// Core 3.10.2: deterministic typed walk, one bounded response window.
// Static facets carry no write capability. Every reused slot is cleared.
FUNCTION "FRK_ConfigRevision" : UDInt
{ S7_Optimized_Access := 'TRUE' }
VERSION : 0.1
VAR_INPUT
    Previous : UDInt;
END_VAR
VAR_TEMP
    Stamp : DTL;
    ResultCode : Int;
    Generation : ULInt;
END_VAR
BEGIN
    #FRK_ConfigRevision := #Previous + 1;
    #ResultCode := RD_SYS_T(OUT => #Stamp);
    IF #ResultCode = 0 THEN
        #Generation := LDT_TO_ULINT(DTL_TO_LDT(#Stamp)) / ULINT#1000000;
        #FRK_ConfigRevision := ULINT_TO_UDINT(#Generation MOD ULINT#4294967296);
    END_IF;
    IF #FRK_ConfigRevision = #Previous THEN #FRK_ConfigRevision := #Previous + 1; END_IF;
    IF #FRK_ConfigRevision = 0 THEN #FRK_ConfigRevision := 1; END_IF;
END_FUNCTION

FUNCTION "FRK_ConfigBegin" : Void
{ S7_Optimized_Access := 'TRUE' }
VERSION : 0.1
VAR_INPUT
    PageIndex : DInt;
    Revision : UDInt;
END_VAR
VAR_IN_OUT
    Cursor : "FRK_ConfigCursor";
    Page : "ST_ConfigPage";
END_VAR
VAR_TEMP
    Index : Int;
END_VAR
BEGIN
    #Cursor.Position := 0;
    #Cursor.First := 0;
    #Page.Revision := #Revision;
    #Page.PageIndex := 0;
    IF #PageIndex >= 0 AND #PageIndex <= 32767 THEN
        #Cursor.First := #PageIndex * 16;
        #Page.PageIndex := DINT_TO_INT(#PageIndex);
    END_IF;
    #Page.PageCount := 1;
    #Page.EntryCount := 0;
    "FRK_UnitScratch".EmptyConfigEntry.ValueType := 1;
    "FRK_UnitScratch".EmptyConfigEntry.Readable := TRUE;
    FOR #Index := 1 TO 16 DO
        #Page.Entries[#Index] := "FRK_UnitScratch".EmptyConfigEntry;
    END_FOR;
END_FUNCTION

FUNCTION "FRK_ConfigAppend" : Void
{ S7_Optimized_Access := 'TRUE' }
VERSION : 0.1
VAR_INPUT
    Scope : String;
    Item : String;
    ValueText : WString;
    ValueType : DInt;
    ReadLevel : DInt;
    Readable : Bool;
END_VAR
VAR_IN_OUT
    Cursor : "FRK_ConfigCursor";
    Page : "ST_ConfigPage";
END_VAR
VAR_TEMP
    Slot : DInt;
END_VAR
BEGIN
    #Slot := #Cursor.Position - #Cursor.First;
    #Cursor.Position := #Cursor.Position + 1;
    IF #Slot < 0 OR #Slot >= 16 THEN RETURN; END_IF;
    #Slot := #Slot + 1;
    #Page.Entries[#Slot].Scope := STRING_TO_WSTRING(#Scope);
    #Page.Entries[#Slot].Item := STRING_TO_WSTRING(#Item);
    #Page.Entries[#Slot].ValueType := #ValueType;
    #Page.Entries[#Slot].ReadLevel := #ReadLevel;
    #Page.Entries[#Slot].Readable := #Readable;
    IF #Readable THEN #Page.Entries[#Slot].ValueText := #ValueText; END_IF;
    #Page.EntryCount := DINT_TO_INT(#Slot);
END_FUNCTION

FUNCTION "FRK_ConfigFinish" : Void
{ S7_Optimized_Access := 'TRUE' }
VERSION : 0.1
VAR_IN_OUT
    Cursor : "FRK_ConfigCursor";
    Page : "ST_ConfigPage";
END_VAR
BEGIN
    #Page.PageCount := DINT_TO_INT((#Cursor.Position + 16 - 1) / 16);
    IF #Page.PageCount < 1 THEN #Page.PageCount := 1; END_IF;
END_FUNCTION

FUNCTION "FRK_ConfigCatalog" : Void
{ S7_Optimized_Access := 'TRUE' }
VERSION : 0.1
VAR_INPUT
    Scope : String;
    Count : Int;
    Catalog : Array[1..12] of "ST_CommandInfo";
    ReadLevel : DInt;
    Readable : Bool;
END_VAR
VAR_IN_OUT
    Cursor : "FRK_ConfigCursor";
    Page : "ST_ConfigPage";
END_VAR
VAR_TEMP
    Index : Int;
    IndexText : String[8];
    Prefix : String[254];
    Item : String[254];
END_VAR
BEGIN
    "FRK_ConfigAppend"(Scope := #Scope, Item := 'CatalogCount', ValueText := STRING_TO_WSTRING(INT_TO_STRING(#Count)), ValueType := 0, ReadLevel := #ReadLevel, Readable := #Readable, Cursor := #Cursor, Page := #Page);
    FOR #Index := 1 TO #Count DO
        IF #Index > 12 THEN EXIT; END_IF;
        #IndexText := INT_TO_STRING(#Index);
        IF #IndexText[1] = '+' THEN #IndexText := DELETE(IN := #IndexText, L := 1, P := 1); END_IF;
        #Prefix := CONCAT(IN1 := 'Catalog/Catalog[', IN2 := #IndexText);
        #Prefix := CONCAT(IN1 := #Prefix, IN2 := ']/');
        #Item := CONCAT(IN1 := #Prefix, IN2 := 'Value');
        "FRK_ConfigAppend"(Scope := #Scope, Item := #Item, ValueText := STRING_TO_WSTRING(DINT_TO_STRING(#Catalog[#Index].Value)), ValueType := 0, ReadLevel := #ReadLevel, Readable := #Readable, Cursor := #Cursor, Page := #Page);
        #Item := CONCAT(IN1 := #Prefix, IN2 := 'Label');
        "FRK_ConfigAppend"(Scope := #Scope, Item := #Item, ValueText := STRING_TO_WSTRING(#Catalog[#Index].Label), ValueType := 1, ReadLevel := #ReadLevel, Readable := #Readable, Cursor := #Cursor, Page := #Page);
        #Item := CONCAT(IN1 := #Prefix, IN2 := 'Style');
        "FRK_ConfigAppend"(Scope := #Scope, Item := #Item, ValueText := STRING_TO_WSTRING(DINT_TO_STRING(#Catalog[#Index].Style)), ValueType := 0, ReadLevel := #ReadLevel, Readable := #Readable, Cursor := #Cursor, Page := #Page);
    END_FOR;
END_FUNCTION

FUNCTION "FRK_ConfigUnit" : Void
{ S7_Optimized_Access := 'TRUE' }
VERSION : 0.1
VAR_INPUT
    Scope : String;
    Policy : Array[0..6] of "ST_ModePolicy";
    ModelCount : Int;
    ReadLevel : DInt;
    Readable : Bool;
END_VAR
VAR_IN_OUT
    Cursor : "FRK_ConfigCursor";
    Page : "ST_ConfigPage";
END_VAR
VAR_TEMP
    Index : Int;
    IndexText : String[8];
    Prefix : String[254];
    Item : String[254];
END_VAR
BEGIN
    "FRK_ConfigAppend"(Scope := #Scope, Item := 'CatalogCount', ValueText := WSTRING#'0', ValueType := 0, ReadLevel := #ReadLevel, Readable := #Readable, Cursor := #Cursor, Page := #Page);
    "FRK_ConfigAppend"(Scope := #Scope, Item := 'AvailableModelCount', ValueText := INT_TO_WSTRING(#ModelCount), ValueType := 0, ReadLevel := #ReadLevel, Readable := #Readable, Cursor := #Cursor, Page := #Page);
    FOR #Index := 0 TO 6 DO
        #IndexText := INT_TO_STRING(#Index);
        IF #IndexText[1] = '+' THEN #IndexText := DELETE(IN := #IndexText, L := 1, P := 1); END_IF;
        #Prefix := CONCAT(IN1 := 'ModePolicy/ModePolicy[', IN2 := #IndexText);
        #Prefix := CONCAT(IN1 := #Prefix, IN2 := ']/');
        #Item := CONCAT(IN1 := #Prefix, IN2 := 'Shield');
        "FRK_ConfigAppend"(Scope := #Scope, Item := #Item, ValueText := STRING_TO_WSTRING(DINT_TO_STRING(#Policy[#Index].Shield)), ValueType := 0, ReadLevel := #ReadLevel, Readable := #Readable, Cursor := #Cursor, Page := #Page);
        #Item := CONCAT(IN1 := #Prefix, IN2 := 'Style');
        "FRK_ConfigAppend"(Scope := #Scope, Item := #Item, ValueText := STRING_TO_WSTRING(DINT_TO_STRING(#Policy[#Index].Style)), ValueType := 0, ReadLevel := #ReadLevel, Readable := #Readable, Cursor := #Cursor, Page := #Page);
    END_FOR;
END_FUNCTION

// Core 8.3: one owning active list / closed ring, with optional event callback.
FUNCTION "FRK_AlarmNotify" : Void
{ S7_Optimized_Access := 'TRUE' }
VERSION : 0.1
VAR_INPUT
    Ev : "ST_AlarmEvent";
END_VAR
VAR_IN_OUT
    AlarmLog : "FRK_AlarmLog";
END_VAR
BEGIN
    RETURN; // No event sink supplied by the composition declaration.
END_FUNCTION

FUNCTION "FRK_AlarmRefresh" : Void
{ S7_Optimized_Access := 'TRUE' }
VERSION : 0.1
VAR_IN_OUT
    AlarmLog : "FRK_AlarmLog";
END_VAR
VAR_TEMP
    Index : Int;
END_VAR
BEGIN
    #AlarmLog.NActive := 0;
    #AlarmLog.Blocking := FALSE;
    FOR #Index := 1 TO 16 DO
        IF #AlarmLog.Active[#Index].State <> 0 THEN
            #AlarmLog.NActive := #AlarmLog.NActive + 1;
            IF #AlarmLog.Active[#Index].ResetClass = 1 THEN #AlarmLog.Blocking := TRUE; END_IF;
        END_IF;
    END_FOR;
END_FUNCTION

FUNCTION "FRK_AlarmBegin" : Void
{ S7_Optimized_Access := 'TRUE' }
VERSION : 0.1
VAR_INPUT
    Startup : Bool;
END_VAR
VAR_IN_OUT
    AlarmLog : "FRK_AlarmLog";
END_VAR
VAR_TEMP
    Index : Int;
END_VAR
BEGIN
    FOR #Index := 1 TO 16 DO
        #AlarmLog.Touched[#Index] := FALSE;
        IF #Startup THEN
            #AlarmLog.Active[#Index] := "FRK_UnitScratch".EmptyEvent;
            #AlarmLog.Automatic[#Index] := FALSE;
            #AlarmLog.ComeMs[#Index] := 0;
        END_IF;
    END_FOR;
    IF #Startup THEN
        FOR #Index := 1 TO 64 DO #AlarmLog.Ring[#Index] := "FRK_UnitScratch".EmptyEvent; END_FOR;
        #AlarmLog.RingHead := 0;
        #AlarmLog.RingUsed := 0;
        #AlarmLog.Truncated := FALSE;
    END_IF;
    "FRK_AlarmRefresh"(AlarmLog := #AlarmLog);
END_FUNCTION

FUNCTION "FRK_AlarmRaise" : Int
{ S7_Optimized_Access := 'TRUE' }
VERSION : 0.1
VAR_INPUT
    Diag : "ST_Diagnostic";
    ResetClass : DInt;
END_VAR
VAR_IN_OUT
    AlarmLog : "FRK_AlarmLog";
END_VAR
VAR_TEMP
    Slot : Int;
    Stamp : DTL;
    ResultCode : Int;
    Rational : "ST_Diagnostic";
END_VAR
BEGIN
    #FRK_AlarmRaise := 0;
    IF #ResetClass < 0 OR #ResetClass > 1
        OR #Diag.Severity < 0 OR #Diag.Severity > 2
        OR #Diag.Category < 0 OR #Diag.Category > 2
        OR #Diag.SourcePath = WSTRING#'' OR #Diag.Description = WSTRING#'' THEN RETURN; END_IF;
    FOR #Slot := 1 TO 16 DO
        IF #AlarmLog.Active[#Slot].State = 0 THEN
            #Rational := #Diag;
            "FRK_Rationalize"(Diag := #Rational);
            #AlarmLog.Active[#Slot] := "FRK_UnitScratch".EmptyEvent;
            #AlarmLog.Active[#Slot].ReasonCode := #Rational.ReasonCode;
            #AlarmLog.Active[#Slot].Description := #Rational.Description;
            #AlarmLog.Active[#Slot].SourcePath := #Rational.SourcePath;
            #AlarmLog.Active[#Slot].IoTag := #Rational.IoTag;
            #AlarmLog.Active[#Slot].IoAddress := #Rational.IoAddress;
            #AlarmLog.Active[#Slot].Severity := #Rational.Severity;
            #AlarmLog.Active[#Slot].Category := #Rational.Category;
            #AlarmLog.Active[#Slot].ResetClass := #ResetClass;
            #AlarmLog.Active[#Slot].State := 1;
            #AlarmLog.ComeMs[#Slot] := "FRK_Clock".NowMs;
            #AlarmLog.Automatic[#Slot] := FALSE;
            #AlarmLog.Touched[#Slot] := FALSE;
            #ResultCode := RD_SYS_T(OUT => #Stamp);
            IF #ResultCode = 0 THEN #AlarmLog.Active[#Slot].ComeAt := DTL_TO_LDT(#Stamp); END_IF;
            // The UTC source has no proven synchronization witness yet.
            #AlarmLog.Active[#Slot].ComeTimeSynchronized := FALSE;
            "FRK_AlarmRefresh"(AlarmLog := #AlarmLog);
            "FRK_AlarmNotify"(AlarmLog := #AlarmLog, Ev := #AlarmLog.Active[#Slot]);
            #FRK_AlarmRaise := #Slot;
            RETURN;
        END_IF;
    END_FOR;
    #AlarmLog.Truncated := TRUE;
END_FUNCTION

FUNCTION "FRK_AlarmClose" : Void
{ S7_Optimized_Access := 'TRUE' }
VERSION : 0.1
VAR_INPUT
    Slot : Int;
END_VAR
VAR_IN_OUT
    AlarmLog : "FRK_AlarmLog";
END_VAR
BEGIN
    IF #Slot < 1 OR #Slot > 16 THEN RETURN; END_IF;
    IF #AlarmLog.Active[#Slot].State = 0 THEN RETURN; END_IF;
    #AlarmLog.Active[#Slot].State := 0;
    IF #AlarmLog.RingHead < 0 OR #AlarmLog.RingHead > 64 THEN #AlarmLog.RingHead := 0; END_IF;
    #AlarmLog.RingHead := (#AlarmLog.RingHead MOD 64) + 1;
    IF #AlarmLog.RingUsed >= 64 THEN #AlarmLog.Truncated := TRUE;
    ELSE #AlarmLog.RingUsed := #AlarmLog.RingUsed + 1; END_IF;
    #AlarmLog.Ring[#AlarmLog.RingHead] := #AlarmLog.Active[#Slot];
    #AlarmLog.Automatic[#Slot] := FALSE;
    "FRK_AlarmRefresh"(AlarmLog := #AlarmLog);
    "FRK_AlarmNotify"(AlarmLog := #AlarmLog, Ev := #AlarmLog.Ring[#AlarmLog.RingHead]);
END_FUNCTION

FUNCTION "FRK_AlarmGone" : Bool
{ S7_Optimized_Access := 'TRUE' }
VERSION : 0.1
VAR_INPUT
    Slot : Int;
END_VAR
VAR_IN_OUT
    AlarmLog : "FRK_AlarmLog";
END_VAR
VAR_TEMP
    Span : UDInt;
    Stamp : DTL;
    ResultCode : Int;
END_VAR
BEGIN
    #FRK_AlarmGone := FALSE;
    IF #Slot < 1 OR #Slot > 16 THEN RETURN; END_IF;
    IF #AlarmLog.Active[#Slot].State <> 1 THEN RETURN; END_IF;
    #ResultCode := RD_SYS_T(OUT => #Stamp);
    IF #ResultCode = 0 THEN #AlarmLog.Active[#Slot].GoneAt := DTL_TO_LDT(#Stamp); END_IF;
    #AlarmLog.Active[#Slot].GoneTimeSynchronized := FALSE;
    #Span := "FRK_Elapsed"(NewMs := "FRK_Clock".NowMs, OldMs := #AlarmLog.ComeMs[#Slot]);
    IF #Span > 2147483647 THEN #Span := 2147483647; END_IF;
    #AlarmLog.Active[#Slot].Duration := DINT_TO_TIME(UDINT_TO_DINT(#Span));
    IF #AlarmLog.Active[#Slot].ResetClass = 0 THEN
        "FRK_AlarmClose"(AlarmLog := #AlarmLog, Slot := #Slot);
    ELSE
        #AlarmLog.Active[#Slot].State := 2;
        #AlarmLog.Automatic[#Slot] := FALSE;
    END_IF;
    #FRK_AlarmGone := TRUE;
END_FUNCTION

FUNCTION "FRK_AlarmOperatorReset" : Void
{ S7_Optimized_Access := 'TRUE' }
VERSION : 0.1
VAR_IN_OUT
    AlarmLog : "FRK_AlarmLog";
END_VAR
VAR_TEMP
    Slot : Int;
    Gone : Bool;
    Stamp : DTL;
    ResultCode : Int;
END_VAR
BEGIN
    FOR #Slot := 1 TO 16 DO
        IF #AlarmLog.Active[#Slot].State <> 0 AND #AlarmLog.Active[#Slot].ResetClass = 1 THEN
            IF #AlarmLog.Active[#Slot].State = 1 THEN #Gone := "FRK_AlarmGone"(AlarmLog := #AlarmLog, Slot := #Slot); END_IF;
            #ResultCode := RD_SYS_T(OUT => #Stamp);
            IF #ResultCode = 0 THEN #AlarmLog.Active[#Slot].ResetAt := DTL_TO_LDT(#Stamp); END_IF;
            #AlarmLog.Active[#Slot].ResetTimeSynchronized := FALSE;
            "FRK_AlarmClose"(AlarmLog := #AlarmLog, Slot := #Slot);
        END_IF;
    END_FOR;
END_FUNCTION

FUNCTION "FRK_AlarmMessage" : Void
{ S7_Optimized_Access := 'TRUE' }
VERSION : 0.1
VAR_INPUT
    Reason : DInt;
    Description : WString;
    SourcePath : WString;
END_VAR
VAR_IN_OUT
    AlarmLog : "FRK_AlarmLog";
END_VAR
VAR_TEMP
    Diag : "ST_Diagnostic";
    Slot : Int;
    Gone : Bool;
END_VAR
BEGIN
    #Diag := "FRK_UnitScratch".EmptyDiagnostic;
    #Diag.ReasonCode := #Reason;
    #Diag.Description := #Description;
    #Diag.SourcePath := #SourcePath;
    #Diag.Severity := 0;
    #Diag.Category := 2;
    #Slot := "FRK_AlarmRaise"(AlarmLog := #AlarmLog, Diag := #Diag, ResetClass := 0);
    IF #Slot > 0 THEN #Gone := "FRK_AlarmGone"(AlarmLog := #AlarmLog, Slot := #Slot); END_IF;
END_FUNCTION

FUNCTION "FRK_AlarmCapture" : Void
{ S7_Optimized_Access := 'TRUE' }
VERSION : 0.1
VAR_IN_OUT
    AlarmLog : "FRK_AlarmLog";
    Core : "FRK_Core";
    Status : "ST_ModuleStatus";
END_VAR
VAR_TEMP
    Slot : Int;
END_VAR
BEGIN
    #Slot := #Core.FaultSlot;
    IF #Slot < 1 OR #Slot > 16 THEN #Slot := 0;
    ELSIF NOT #AlarmLog.Automatic[#Slot] OR #AlarmLog.Active[#Slot].State <> 1
        OR #AlarmLog.Active[#Slot].SourcePath <> #Status.Diagnostic.SourcePath
        OR #AlarmLog.Active[#Slot].ReasonCode <> #Status.Diagnostic.ReasonCode
        OR #AlarmLog.Active[#Slot].Description <> #Status.Diagnostic.Description THEN #Slot := 0; END_IF;
    IF #Core.Exec = 3 THEN
        IF #Slot = 0 THEN
            // Adopted first-outs share one active occurrence within this log.
            FOR #Slot := 1 TO 16 DO
                IF #AlarmLog.Automatic[#Slot] AND #AlarmLog.Active[#Slot].State = 1
                    AND #AlarmLog.Active[#Slot].SourcePath = #Status.Diagnostic.SourcePath
                    AND #AlarmLog.Active[#Slot].ReasonCode = #Status.Diagnostic.ReasonCode
                    AND #AlarmLog.Active[#Slot].Description = #Status.Diagnostic.Description THEN EXIT; END_IF;
            END_FOR;
            IF #Slot > 16 THEN #Slot := "FRK_AlarmRaise"(AlarmLog := #AlarmLog, Diag := #Status.Diagnostic, ResetClass := 1); END_IF;
        END_IF;
        IF #Slot > 0 THEN #AlarmLog.Automatic[#Slot] := TRUE; #AlarmLog.Touched[#Slot] := TRUE; END_IF;
        #Core.FaultSlot := #Slot;
    ELSE
        #Core.FaultSlot := 0;
    END_IF;
END_FUNCTION

FUNCTION "FRK_AlarmEnd" : Void
{ S7_Optimized_Access := 'TRUE' }
VERSION : 0.1
VAR_IN_OUT
    AlarmLog : "FRK_AlarmLog";
END_VAR
VAR_TEMP
    Slot : Int;
    Gone : Bool;
END_VAR
BEGIN
    FOR #Slot := 1 TO 16 DO
        IF #AlarmLog.Automatic[#Slot] AND NOT #AlarmLog.Touched[#Slot] THEN #Gone := "FRK_AlarmGone"(AlarmLog := #AlarmLog, Slot := #Slot); END_IF;
    END_FOR;
END_FUNCTION

FUNCTION "FRK_AlarmTreeBlocking" : Bool
{ S7_Optimized_Access := 'TRUE' }
VERSION : 0.1
VAR_INPUT
    Owner : DInt;
END_VAR
VAR_TEMP
    Index : DInt;
    Ancestor : DInt;
    Depth : DInt;
END_VAR
BEGIN
    #FRK_AlarmTreeBlocking := TRUE;
    IF "FRK_Registry".Fault OR #Owner < 1 OR #Owner > "FRK_Registry".Count OR "FRK_Registry".Count > 32 THEN RETURN; END_IF;
    FOR #Index := 1 TO "FRK_Registry".Count DO
        IF "FRK_Registry".Rows[#Index].AlarmBlocking THEN
            #Ancestor := #Index;
            FOR #Depth := 1 TO 32 DO
                IF #Ancestor = #Owner THEN RETURN; END_IF;
                IF #Ancestor = 0 THEN EXIT; END_IF;
                IF #Ancestor < 1 OR #Ancestor > "FRK_Registry".Count THEN RETURN; END_IF;
                #Ancestor := "FRK_Registry".Rows[#Ancestor].Parent;
            END_FOR;
            IF #Depth > 32 AND #Ancestor <> 0 THEN RETURN; END_IF;
        END_IF;
    END_FOR;
    #FRK_AlarmTreeBlocking := FALSE;
END_FUNCTION

// Core section 7.7 prototype: volatile provider injection and independent root sessions.
// User records are salted Core-compatible hashes, never commissioning plaintext.
FUNCTION "FRK_Sha256Pin" : Bool
{ S7_Optimized_Access := 'TRUE' }
VERSION : 0.1
VAR_INPUT
    Size : DInt;
END_VAR
VAR_IN_OUT
    Data : Array[0..47] of Byte;
    Digest : Array[0..31] of Byte;
END_VAR
VAR_TEMP
    BlockBytes : Array[0..63] of Byte;
    Words : Array[0..63] of DWord;
    Hash : Array[0..7] of DWord;
    Index : DInt;
    A : DWord;
    B : DWord;
    C : DWord;
    D : DWord;
    E : DWord;
    F : DWord;
    G : DWord;
    H : DWord;
    S0 : DWord;
    S1 : DWord;
    T1 : DWord;
    T2 : DWord;
    K : Array[0..63] of DWord;
END_VAR
BEGIN
    #FRK_Sha256Pin := FALSE;
    #K[0] := DWORD#16#428A2F98;
    #K[1] := DWORD#16#71374491;
    #K[2] := DWORD#16#B5C0FBCF;
    #K[3] := DWORD#16#E9B5DBA5;
    #K[4] := DWORD#16#3956C25B;
    #K[5] := DWORD#16#59F111F1;
    #K[6] := DWORD#16#923F82A4;
    #K[7] := DWORD#16#AB1C5ED5;
    #K[8] := DWORD#16#D807AA98;
    #K[9] := DWORD#16#12835B01;
    #K[10] := DWORD#16#243185BE;
    #K[11] := DWORD#16#550C7DC3;
    #K[12] := DWORD#16#72BE5D74;
    #K[13] := DWORD#16#80DEB1FE;
    #K[14] := DWORD#16#9BDC06A7;
    #K[15] := DWORD#16#C19BF174;
    #K[16] := DWORD#16#E49B69C1;
    #K[17] := DWORD#16#EFBE4786;
    #K[18] := DWORD#16#0FC19DC6;
    #K[19] := DWORD#16#240CA1CC;
    #K[20] := DWORD#16#2DE92C6F;
    #K[21] := DWORD#16#4A7484AA;
    #K[22] := DWORD#16#5CB0A9DC;
    #K[23] := DWORD#16#76F988DA;
    #K[24] := DWORD#16#983E5152;
    #K[25] := DWORD#16#A831C66D;
    #K[26] := DWORD#16#B00327C8;
    #K[27] := DWORD#16#BF597FC7;
    #K[28] := DWORD#16#C6E00BF3;
    #K[29] := DWORD#16#D5A79147;
    #K[30] := DWORD#16#06CA6351;
    #K[31] := DWORD#16#14292967;
    #K[32] := DWORD#16#27B70A85;
    #K[33] := DWORD#16#2E1B2138;
    #K[34] := DWORD#16#4D2C6DFC;
    #K[35] := DWORD#16#53380D13;
    #K[36] := DWORD#16#650A7354;
    #K[37] := DWORD#16#766A0ABB;
    #K[38] := DWORD#16#81C2C92E;
    #K[39] := DWORD#16#92722C85;
    #K[40] := DWORD#16#A2BFE8A1;
    #K[41] := DWORD#16#A81A664B;
    #K[42] := DWORD#16#C24B8B70;
    #K[43] := DWORD#16#C76C51A3;
    #K[44] := DWORD#16#D192E819;
    #K[45] := DWORD#16#D6990624;
    #K[46] := DWORD#16#F40E3585;
    #K[47] := DWORD#16#106AA070;
    #K[48] := DWORD#16#19A4C116;
    #K[49] := DWORD#16#1E376C08;
    #K[50] := DWORD#16#2748774C;
    #K[51] := DWORD#16#34B0BCB5;
    #K[52] := DWORD#16#391C0CB3;
    #K[53] := DWORD#16#4ED8AA4A;
    #K[54] := DWORD#16#5B9CCA4F;
    #K[55] := DWORD#16#682E6FF3;
    #K[56] := DWORD#16#748F82EE;
    #K[57] := DWORD#16#78A5636F;
    #K[58] := DWORD#16#84C87814;
    #K[59] := DWORD#16#8CC70208;
    #K[60] := DWORD#16#90BEFFFA;
    #K[61] := DWORD#16#A4506CEB;
    #K[62] := DWORD#16#BEF9A3F7;
    #K[63] := DWORD#16#C67178F2;
    FOR #Index := 0 TO 31 DO #Digest[#Index] := 0; END_FOR;
    IF #Size < 0 OR #Size > 48 THEN RETURN; END_IF;
    // Authentication messages fit exactly one SHA-256 block.
    FOR #Index := 0 TO 63 DO #BlockBytes[#Index] := 0; END_FOR;
    FOR #Index := 0 TO #Size - 1 DO #BlockBytes[#Index] := #Data[#Index]; END_FOR;
    #BlockBytes[#Size] := BYTE#16#80;
    #BlockBytes[62] := DWORD_TO_BYTE(SHR(IN := DINT_TO_DWORD(#Size * 8), N := 8));
    #BlockBytes[63] := DINT_TO_BYTE(#Size * 8);
    #Hash[0] := DWORD#16#6A09E667;
    #Hash[1] := DWORD#16#BB67AE85;
    #Hash[2] := DWORD#16#3C6EF372;
    #Hash[3] := DWORD#16#A54FF53A;
    #Hash[4] := DWORD#16#510E527F;
    #Hash[5] := DWORD#16#9B05688C;
    #Hash[6] := DWORD#16#1F83D9AB;
    #Hash[7] := DWORD#16#5BE0CD19;
    FOR #Index := 0 TO 15 DO
        #Words[#Index] := SHL(IN := BYTE_TO_DWORD(#BlockBytes[4 * #Index]), N := 24)
            OR SHL(IN := BYTE_TO_DWORD(#BlockBytes[4 * #Index + 1]), N := 16)
            OR SHL(IN := BYTE_TO_DWORD(#BlockBytes[4 * #Index + 2]), N := 8)
            OR BYTE_TO_DWORD(#BlockBytes[4 * #Index + 3]);
    END_FOR;
    FOR #Index := 16 TO 63 DO
        #S0 := ROR(IN := #Words[#Index-15], N := 7) XOR ROR(IN := #Words[#Index-15], N := 18) XOR SHR(IN := #Words[#Index-15], N := 3);
        #S1 := ROR(IN := #Words[#Index-2], N := 17) XOR ROR(IN := #Words[#Index-2], N := 19) XOR SHR(IN := #Words[#Index-2], N := 10);
        #Words[#Index] := UDINT_TO_DWORD(ULINT_TO_UDINT(UDINT_TO_ULINT(DWORD_TO_UDINT(#Words[#Index-16])) + UDINT_TO_ULINT(DWORD_TO_UDINT(#S0)) + UDINT_TO_ULINT(DWORD_TO_UDINT(#Words[#Index-7])) + UDINT_TO_ULINT(DWORD_TO_UDINT(#S1))));
    END_FOR;
    #A := #Hash[0]; #B := #Hash[1]; #C := #Hash[2]; #D := #Hash[3];
    #E := #Hash[4]; #F := #Hash[5]; #G := #Hash[6]; #H := #Hash[7];
    FOR #Index := 0 TO 63 DO
        #S1 := ROR(IN := #E, N := 6) XOR ROR(IN := #E, N := 11) XOR ROR(IN := #E, N := 25);
        #T1 := UDINT_TO_DWORD(ULINT_TO_UDINT(UDINT_TO_ULINT(DWORD_TO_UDINT(#H)) + UDINT_TO_ULINT(DWORD_TO_UDINT(#S1)) + UDINT_TO_ULINT(DWORD_TO_UDINT((#E AND #F) XOR ((NOT #E) AND #G))) + UDINT_TO_ULINT(DWORD_TO_UDINT(#K[#Index])) + UDINT_TO_ULINT(DWORD_TO_UDINT(#Words[#Index]))));
        #S0 := ROR(IN := #A, N := 2) XOR ROR(IN := #A, N := 13) XOR ROR(IN := #A, N := 22);
        #T2 := UDINT_TO_DWORD(ULINT_TO_UDINT(UDINT_TO_ULINT(DWORD_TO_UDINT(#S0)) + UDINT_TO_ULINT(DWORD_TO_UDINT((#A AND #B) XOR (#A AND #C) XOR (#B AND #C)))));
        #H := #G; #G := #F; #F := #E;
        #E := UDINT_TO_DWORD(ULINT_TO_UDINT(UDINT_TO_ULINT(DWORD_TO_UDINT(#D)) + UDINT_TO_ULINT(DWORD_TO_UDINT(#T1))));
        #D := #C; #C := #B; #B := #A;
        #A := UDINT_TO_DWORD(ULINT_TO_UDINT(UDINT_TO_ULINT(DWORD_TO_UDINT(#T1)) + UDINT_TO_ULINT(DWORD_TO_UDINT(#T2))));
    END_FOR;
    #Words[0] := #A; #Words[1] := #B; #Words[2] := #C; #Words[3] := #D;
    #Words[4] := #E; #Words[5] := #F; #Words[6] := #G; #Words[7] := #H;
    FOR #Index := 0 TO 7 DO
        #Hash[#Index] := UDINT_TO_DWORD(ULINT_TO_UDINT(UDINT_TO_ULINT(DWORD_TO_UDINT(#Hash[#Index])) + UDINT_TO_ULINT(DWORD_TO_UDINT(#Words[#Index]))));
        #Digest[4 * #Index] := DWORD_TO_BYTE(SHR(IN := #Hash[#Index], N := 24));
        #Digest[4 * #Index + 1] := DWORD_TO_BYTE(SHR(IN := #Hash[#Index], N := 16));
        #Digest[4 * #Index + 2] := DWORD_TO_BYTE(SHR(IN := #Hash[#Index], N := 8));
        #Digest[4 * #Index + 3] := DWORD_TO_BYTE(#Hash[#Index]);
    END_FOR;
    FOR #Index := 0 TO 63 DO #BlockBytes[#Index] := 0; #Words[#Index] := 0; END_FOR;
    #FRK_Sha256Pin := TRUE;
END_FUNCTION

FUNCTION "FRK_AccessCancel" : Void
{ S7_Optimized_Access := 'TRUE' }
VERSION : 0.1
VAR_IN_OUT
    Access : "FRK_Access";
END_VAR
VAR_TEMP
    Index : DInt;
END_VAR
BEGIN
    #Access.LoginBusy := FALSE;
    #Access.CandidateUser := '';
    #Access.CandidateLevel := 0;
    #Access.Round := 0;
    FOR #Index := 0 TO 15 DO #Access.Salt[#Index] := 0; END_FOR;
    FOR #Index := 0 TO 31 DO #Access.Digest[#Index] := 0; #Access.Expected[#Index] := 0; END_FOR;
END_FUNCTION

FUNCTION "FRK_AccessLogout" : Void
{ S7_Optimized_Access := 'TRUE' }
VERSION : 0.1
VAR_IN_OUT
    Access : "FRK_Access";
END_VAR
BEGIN
    "FRK_AccessCancel"(Access := #Access);
    "FRK_AccessDropSession"(Access := #Access);
END_FUNCTION

FUNCTION "FRK_AccessDropSession" : Void
{ S7_Optimized_Access := 'TRUE' }
VERSION : 0.1
VAR_IN_OUT
    Access : "FRK_Access";
END_VAR
BEGIN
    #Access.CurrentLevel := 0;
    #Access.CurrentUser := '';
    #Access.LoginFailed := FALSE;
    #Access.SessionGeneration := "FRK_AccessNext"(Previous := #Access.SessionGeneration);
END_FUNCTION

FUNCTION "FRK_AccessNext" : UDInt
{ S7_Optimized_Access := 'TRUE' }
VERSION : 0.1
VAR_INPUT
    Previous : UDInt;
END_VAR
BEGIN
    IF #Previous = UDINT#4294967295 THEN #FRK_AccessNext := 1; ELSE #FRK_AccessNext := #Previous + 1; END_IF;
END_FUNCTION

FUNCTION "FRK_AccessLogin" : Void
{ S7_Optimized_Access := 'TRUE' }
VERSION : 0.1
VAR_INPUT
    User : String;
    Secret : String;
    Sequence : UDInt;
END_VAR
VAR_IN_OUT
    Access : "FRK_Access";
END_VAR
VAR_TEMP
    Data : Array[0..47] of Byte;
    Index : DInt;
    Slot : DInt;
    Size : Int;
    HashOk : Bool;
END_VAR
BEGIN
    "FRK_AccessCancel"(Access := #Access);
    #Access.LoginFailed := FALSE;
    #Access.LoginSequence := #Sequence;
    #Access.LoginSince := "FRK_Clock".NowMs;
    #Access.LoginTimeoutMs := 6000;
    #Access.CandidateUser := #User;
    // Unknown users execute the same bounded work with a dummy salt/digest.
    IF #Access.ProviderEnabled AND "FRK_LocalUsers".Count >= 0 AND "FRK_LocalUsers".Count <= 16 THEN
        FOR #Slot := 1 TO "FRK_LocalUsers".Count DO
            IF #User <> '' AND "FRK_LocalUsers".Rows[#Slot].User = #User THEN
                IF "FRK_LocalUsers".Rows[#Slot].Level >= 1 AND "FRK_LocalUsers".Rows[#Slot].Level <= 4 THEN
                    #Access.CandidateLevel := "FRK_LocalUsers".Rows[#Slot].Level;
                    #Access.Salt := "FRK_LocalUsers".Rows[#Slot].Salt;
                    #Access.Expected := "FRK_LocalUsers".Rows[#Slot].PinHash;
                END_IF;
                EXIT;
            END_IF;
        END_FOR;
    END_IF;
    FOR #Index := 0 TO 47 DO #Data[#Index] := 0; END_FOR;
    FOR #Index := 0 TO 15 DO #Data[#Index] := #Access.Salt[#Index]; END_FOR;
    #Size := LEN(#Secret);
    IF #Size > 32 THEN #Size := 0; #Access.CandidateLevel := 0; END_IF;
    FOR #Index := 1 TO #Size DO #Data[15 + #Index] := CHAR_TO_BYTE(#Secret[#Index]); END_FOR;
    #HashOk := "FRK_Sha256Pin"(Data := #Data, Size := 16 + INT_TO_DINT(#Size), Digest := #Access.Digest);
    FOR #Index := 0 TO 47 DO #Data[#Index] := 0; END_FOR;
    #Access.LoginBusy := #HashOk;
END_FUNCTION

FUNCTION "FRK_AccessAudit" : Void
{ S7_Optimized_Access := 'TRUE' }
VERSION : 0.1
VAR_INPUT
    What : WString;
    Who : String;
    SourcePath : WString;
END_VAR
VAR_IN_OUT
    AlarmLog : "FRK_AlarmLog";
END_VAR
VAR_TEMP
    Description : WString[480];
END_VAR
BEGIN
    #Description := CONCAT(IN1 := #What, IN2 := WSTRING#': ');
    #Description := CONCAT(IN1 := #Description, IN2 := STRING_TO_WSTRING(#Who));
    "FRK_AlarmMessage"(AlarmLog := #AlarmLog, Reason := 0, Description := #Description, SourcePath := #SourcePath);
END_FUNCTION

FUNCTION "FRK_AccessCyclic" : Void
{ S7_Optimized_Access := 'TRUE' }
VERSION : 0.1
VAR_INPUT
    Startup : Bool;
    SourcePath : WString;
END_VAR
VAR_IN_OUT
    Access : "FRK_Access";
    AlarmLog : "FRK_AlarmLog";
    Revision : UDInt;
END_VAR
VAR_TEMP
    Data : Array[0..47] of Byte;
    Index : DInt;
    Difference : Byte;
    HashOk : Bool;
END_VAR
BEGIN
    #Access.LoginTimeoutMs := 6000;
    IF #Startup THEN
        "FRK_AccessLogout"(Access := #Access);
        #Access.LoginResultSequence := 0;
    END_IF;
    IF #Access.CurrentLevel > 0 AND #Access.Policy.SessionTimeout > T#0ms THEN
        IF "FRK_Elapsed"(NewMs := "FRK_Clock".NowMs, OldMs := #Access.LastActivity) >= DINT_TO_UDINT(TIME_TO_DINT(#Access.Policy.SessionTimeout)) THEN
            "FRK_AccessAudit"(AlarmLog := #AlarmLog, What := WSTRING#'std.audit.autoLogout', Who := #Access.CurrentUser, SourcePath := #SourcePath);
            // Expiring the old session does not discard a separately committed
            // credential attempt. Explicit logout cancels both.
            "FRK_AccessDropSession"(Access := #Access);
            #Revision := "FRK_ConfigRevision"(Previous := #Revision);
        END_IF;
    END_IF;
    IF NOT #Access.LoginBusy THEN RETURN; END_IF;
    // One compression per active scan; never run all PIN rounds in one scan.
    FOR #Index := 0 TO 31 DO #Data[#Index] := #Access.Digest[#Index]; END_FOR;
    FOR #Index := 0 TO 15 DO #Data[32 + #Index] := #Access.Salt[#Index]; END_FOR;
    #HashOk := "FRK_Sha256Pin"(Data := #Data, Size := 48, Digest := #Access.Digest);
    FOR #Index := 0 TO 47 DO #Data[#Index] := 0; END_FOR;
    #Access.Round := #Access.Round + 1;
    IF NOT #HashOk OR "FRK_Elapsed"(NewMs := "FRK_Clock".NowMs, OldMs := #Access.LoginSince) >= #Access.LoginTimeoutMs THEN
        #Access.CandidateLevel := 0;
    ELSIF #Access.Round < 256 THEN RETURN;
    END_IF;
    #Difference := 0;
    FOR #Index := 0 TO 31 DO #Difference := #Difference OR (#Access.Digest[#Index] XOR #Access.Expected[#Index]); END_FOR;
    #Access.LoginFailed := #Difference <> 0 OR #Access.CandidateLevel = 0 OR NOT #Access.ProviderEnabled;
    IF #Access.LoginFailed THEN
        "FRK_AccessAudit"(AlarmLog := #AlarmLog, What := WSTRING#'std.audit.loginFailed', Who := #Access.CandidateUser, SourcePath := #SourcePath);
    ELSE
        #Access.CurrentUser := #Access.CandidateUser;
        #Access.CurrentLevel := #Access.CandidateLevel;
        #Access.LastActivity := "FRK_Clock".NowMs;
        #Access.SessionGeneration := "FRK_AccessNext"(Previous := #Access.SessionGeneration);
        #Revision := "FRK_ConfigRevision"(Previous := #Revision);
        "FRK_AccessAudit"(AlarmLog := #AlarmLog, What := WSTRING#'std.audit.login', Who := #Access.CurrentUser, SourcePath := #SourcePath);
    END_IF;
    #Access.LoginResultSequence := #Access.LoginSequence;
    "FRK_AccessCancel"(Access := #Access);
END_FUNCTION

FUNCTION "FRK_AccessFinish" : Void
{ S7_Optimized_Access := 'TRUE' }
VERSION : 0.1
VAR_INPUT
    Unit : "FRK_Unit";
    Response : "ST_HmiResponse";
    SourcePath : WString;
END_VAR
VAR_IN_OUT
    Access : "FRK_Access";
    AlarmLog : "FRK_AlarmLog";
    Revision : UDInt;
END_VAR
VAR_TEMP
    What : WString[160];
    AuditPath : WString[255];
END_VAR
BEGIN
    IF NOT #Unit.RequestPending THEN RETURN; END_IF;
    CASE #Unit.Request.Kind OF
        23, 15,
        16, 17,
        1: RETURN;
        2:
            "FRK_AccessAudit"(AlarmLog := #AlarmLog, What := WSTRING#'std.audit.logout', Who := #Unit.RequestUser, SourcePath := #SourcePath);
            #Revision := "FRK_ConfigRevision"(Previous := #Revision);
            RETURN;
        ELSE #What := WSTRING#'std.audit.accessDenied';
    END_CASE;
    IF #Response.Accepted THEN
        #What := WSTRING#'std.audit.operatorAction';
        IF #Access.CurrentLevel > 0 THEN #Access.LastActivity := "FRK_Clock".NowMs; END_IF;
        IF #Unit.Request.Kind = 24 THEN #Revision := "FRK_ConfigRevision"(Previous := #Revision); END_IF;
    END_IF;
    #AuditPath := #SourcePath;
    IF #Unit.Request.Kind = 11 THEN
        IF #Response.Accepted THEN #AuditPath := #Unit.Request.TargetPath; END_IF;
        IF #Response.Accepted THEN #What := WSTRING#'std.audit.manualCommandAccepted'; ELSE #What := WSTRING#'std.audit.manualCommandRejected'; END_IF;
    END_IF;
    #What := CONCAT(IN1 := #What, IN2 := WSTRING#' kind=');
    #What := CONCAT(IN1 := #What, IN2 := DINT_TO_WSTRING(#Unit.Request.Kind));
    #What := CONCAT(IN1 := #What, IN2 := WSTRING#' value=');
    #What := CONCAT(IN1 := #What, IN2 := DINT_TO_WSTRING(#Unit.Request.IntValue));
    "FRK_AccessAudit"(AlarmLog := #AlarmLog, What := #What, Who := #Unit.RequestUser, SourcePath := #AuditPath);
END_FUNCTION

// Shared Unit services v0.1: operation authority, mailbox, modes and local carrier.
FUNCTION "FRK_UnitPrepare" : Void
{ S7_Optimized_Access := 'TRUE' }
VERSION : 0.1
VAR_INPUT
    Startup : Bool;
    InitialMode : DInt;
END_VAR
VAR_IN_OUT
    Core : "FRK_Core";
    Unit : "FRK_Unit";
    Policy : Array[0..6] of "ST_ModePolicy";
    Request : "ST_HmiRequest";
    Response : "ST_HmiResponse";
END_VAR
VAR_TEMP
    Index : DInt;
END_VAR
BEGIN
    #Core.EvModeExit := FALSE;
    #Core.EvModeChanged := FALSE;
    IF NOT #Unit.Initialized THEN
        #Unit.Initialized := TRUE;
        #Unit.Permit := TRUE;
        FOR #Index := 0 TO 7-1 DO
            #Policy[#Index].Shield := 1;
            #Policy[#Index].Style := 1;
        END_FOR;
        #Policy[0].Style := 0;
        #Policy[2].Shield := 0;
        #Policy[1].Shield := 0;
        #Policy[3].Shield := 2;
        #Policy[4].Shield := 2;
        #Unit.Mode := #InitialMode;
    END_IF;
    IF #Startup THEN
        #Unit.EvReset := FALSE;
        #Unit.Mode := #InitialMode;
        #Unit.RunReq := FALSE;
        #Unit.AbortReq := #Core.Exec = 1;
        #Unit.StopReq := FALSE;
        #Unit.ModePending := FALSE;
        #Unit.FollowStart := FALSE;
        #Unit.CascadePending := FALSE;
        #Unit.ReleaseChildren := TRUE;
        #Unit.Clearing := TRUE;
        // Consume the restart boundary without executing a transported request.
        #Unit.SeenSequence := #Request.Sequence;
        #Unit.RequestPending := FALSE;
        #Request.Secret := '';
        #Response.Accepted := FALSE;
        #Response.Diagnostic := WSTRING#'std.error.hmiRequestRejected';
        #Response.AckSequence := #Unit.SeenSequence;
    END_IF;
    IF #Core.ReleasePending THEN
        #Unit.FollowStart := FALSE;
        // An incoming parent mode/reset operation is already queued for this scan.
        // Preserve its cascade while cancelling the old command.
        #Unit.RunReq := FALSE;
        #Unit.AbortReq := TRUE;
        #Unit.ReleaseChildren := TRUE;
        #Unit.Clearing := TRUE;
    END_IF;
END_FUNCTION

FUNCTION "FRK_UnitSetLocalCarrier" : Void
{ S7_Optimized_Access := 'TRUE' }
VERSION : 0.1
VAR_INPUT
    Index : DInt;
END_VAR
VAR_IN_OUT
    Unit : "FRK_Unit";
END_VAR
BEGIN
    #Unit.CarrierIndex := 0;
    IF #Index < 1 OR #Index > 32 THEN RETURN; END_IF;
    "FRK_Carriers".Slots[#Index].Enabled := TRUE;
    "FRK_Carriers".Slots[#Index].Kind := 2;
    #Unit.CarrierIndex := #Index;
END_FUNCTION

FUNCTION "FRK_PartEvent" : Void
{ S7_Optimized_Access := 'TRUE' }
VERSION : 0.1
VAR_INPUT
    Reason : DInt;
    Uid : String;
    SourcePath : String;
END_VAR
VAR_IN_OUT
    AlarmLog : "FRK_AlarmLog";
END_VAR
VAR_TEMP
    Description : WString[255];
END_VAR
BEGIN
    CASE #Reason OF
        2024: #Description := WSTRING#'std.event.partReceived: ';
        2025: #Description := WSTRING#'std.event.partProcessingStarted: ';
        2026: #Description := WSTRING#'std.event.partProcessed: ';
        2027: #Description := WSTRING#'std.event.partAborted: ';
        ELSE #Description := WSTRING#'';
    END_CASE;
    #Description := CONCAT(IN1 := #Description, IN2 := STRING_TO_WSTRING(#Uid));
    "FRK_AlarmMessage"(AlarmLog := #AlarmLog, Reason := #Reason, Description := #Description, SourcePath := STRING_TO_WSTRING(#SourcePath));
END_FUNCTION

FUNCTION "FRK_PartReceived" : Bool
{ S7_Optimized_Access := 'TRUE' }
VERSION : 0.1
VAR_IN_OUT
    Core : "FRK_Core";
    Unit : "FRK_Unit";
    Status : "ST_ModuleStatus";
    Part : "ST_PartContext";
    AlarmLog : "FRK_AlarmLog";
END_VAR
VAR_TEMP
    Index : DInt;
    Uid : String[64];
    ResultIndex : DInt;
END_VAR
BEGIN
    #FRK_PartReceived := FALSE;
    #Index := #Unit.CarrierIndex;
    IF #Index = 0 THEN RETURN; END_IF;
    IF #Index < 1 OR #Index > 32 THEN
        "FRK_Fault"(Core := #Core, Status := #Status, ReasonCode := 2020, Description := WSTRING#'std.error.partCarrierReadFailed');
        RETURN;
    END_IF;
    IF NOT "FRK_Carriers".Slots[#Index].Enabled OR "FRK_Carriers".Slots[#Index].Kind <> 2 OR "FRK_Carriers".Slots[#Index].Serial = UDINT#4294967295 THEN
        "FRK_Fault"(Core := #Core, Status := #Status, ReasonCode := 2020, Description := WSTRING#'std.error.partCarrierReadFailed');
        RETURN;
    END_IF;
    "FRK_Carriers".Slots[#Index].Serial := "FRK_Carriers".Slots[#Index].Serial + 1;
    #Uid := CONCAT(IN1 := 'FRK-', IN2 := DINT_TO_STRING(#Index));
    #Uid := CONCAT(IN1 := #Uid, IN2 := '-');
    #Uid := CONCAT(IN1 := #Uid, IN2 := UDINT_TO_STRING("FRK_Carriers".Slots[#Index].Serial));
    #Part.Uid := #Uid;
    #Part.Present := TRUE;
    #Part.CarrierKind := 2;
    #Part.Result.Verdict := 0;
    #Part.Result.ReasonCode := 0;
    #Part.Result.StationPath := STRING_TO_WSTRING(#Status.Name);
    #Part.Result.Stamp := LDT#1970-01-01-00:00:00.000000000;
    #Part.Result.TimeSynchronized := FALSE;
    FOR #ResultIndex := 1 TO 32 DO #Part.Result.Records[#ResultIndex].Name := ''; END_FOR;
    FOR #ResultIndex := 1 TO 8 DO #Part.Parents[#ResultIndex] := ''; END_FOR;
    "FRK_Carriers".Slots[#Index].Context := #Part;
    "FRK_PartEvent"(AlarmLog := #AlarmLog, Reason := 2024, Uid := #Part.Uid, SourcePath := #Status.Name);
    #FRK_PartReceived := TRUE;
END_FUNCTION

FUNCTION "FRK_PartStarted" : Void
{ S7_Optimized_Access := 'TRUE' }
VERSION : 0.1
VAR_IN_OUT
    Unit : "FRK_Unit";
    Status : "ST_ModuleStatus";
    Part : "ST_PartContext";
    AlarmLog : "FRK_AlarmLog";
END_VAR
BEGIN
    IF #Unit.CarrierIndex = 0 OR NOT #Part.Present THEN RETURN; END_IF;
    "FRK_PartEvent"(AlarmLog := #AlarmLog, Reason := 2025, Uid := #Part.Uid, SourcePath := #Status.Name);
END_FUNCTION

FUNCTION "FRK_PartProcessed" : Bool
{ S7_Optimized_Access := 'TRUE' }
VERSION : 0.1
VAR_INPUT
    Verdict : DInt;
    Reason : DInt;
END_VAR
VAR_IN_OUT
    Core : "FRK_Core";
    Unit : "FRK_Unit";
    Status : "ST_ModuleStatus";
    Part : "ST_PartContext";
    AlarmLog : "FRK_AlarmLog";
END_VAR
VAR_TEMP
    Index : DInt;
    Stamp : DTL;
    ResultCode : Int;
END_VAR
BEGIN
    #FRK_PartProcessed := FALSE;
    #Index := #Unit.CarrierIndex;
    IF #Index = 0 OR NOT #Part.Present THEN RETURN; END_IF;
    IF #Verdict < 1 OR #Verdict > 3 OR (#Verdict = 2 AND #Reason = 0) THEN
        "FRK_Fault"(Core := #Core, Status := #Status, ReasonCode := 2023, Description := WSTRING#'std.error.nokReasonRequired');
        RETURN;
    END_IF;
    IF #Index < 1 OR #Index > 32 THEN
        "FRK_Fault"(Core := #Core, Status := #Status, ReasonCode := 2021, Description := WSTRING#'std.error.partCarrierWriteFailed');
        RETURN;
    END_IF;
    IF NOT "FRK_Carriers".Slots[#Index].Enabled THEN
        "FRK_Fault"(Core := #Core, Status := #Status, ReasonCode := 2021, Description := WSTRING#'std.error.partCarrierWriteFailed');
        RETURN;
    END_IF;
    IF #Part.Uid <> "FRK_Carriers".Slots[#Index].Context.Uid THEN
        "FRK_Fault"(Core := #Core, Status := #Status, ReasonCode := 2022, Description := WSTRING#'std.error.partCarrierReadFailed');
        RETURN;
    END_IF;
    #Part.Result.Verdict := #Verdict;
    #Part.Result.ReasonCode := #Reason;
    #Part.Result.StationPath := STRING_TO_WSTRING(#Status.Name);
    #Part.Result.TimeSynchronized := FALSE;
    #ResultCode := RD_SYS_T(OUT => #Stamp);
    IF #ResultCode = 0 THEN #Part.Result.Stamp := DTL_TO_LDT(#Stamp); END_IF;
    "FRK_Carriers".Slots[#Index].Written := #Part;
    IF "FRK_Carriers".Slots[#Index].Writes < UDINT#4294967295 THEN "FRK_Carriers".Slots[#Index].Writes := "FRK_Carriers".Slots[#Index].Writes + 1; END_IF;
    CASE #Verdict OF
        1: IF #Unit.Good < UDINT#4294967295 THEN #Unit.Good := #Unit.Good + 1; END_IF;
        2: IF #Unit.Nok < UDINT#4294967295 THEN #Unit.Nok := #Unit.Nok + 1; END_IF; #Unit.NokReason := #Reason;
        3: IF #Unit.Rework < UDINT#4294967295 THEN #Unit.Rework := #Unit.Rework + 1; END_IF;
        ELSE RETURN;
    END_CASE;
    // The provider result is written before publishing EVENT_PART_PROCESSED.
    "FRK_PartEvent"(AlarmLog := #AlarmLog, Reason := 2026, Uid := #Part.Uid, SourcePath := #Status.Name);
    #Part.Present := FALSE;
    #FRK_PartProcessed := TRUE;
END_FUNCTION

FUNCTION "FRK_PartAborted" : Void
{ S7_Optimized_Access := 'TRUE' }
VERSION : 0.1
VAR_IN_OUT
    Core : "FRK_Core";
    Unit : "FRK_Unit";
    Status : "ST_ModuleStatus";
    Part : "ST_PartContext";
    AlarmLog : "FRK_AlarmLog";
END_VAR
BEGIN
    IF #Unit.CarrierIndex = 0 OR NOT #Part.Present THEN RETURN; END_IF;
    #Part.Result.Verdict := 0;
    IF #Core.Exec = 3 AND #Part.Result.ReasonCode = 0 THEN #Part.Result.ReasonCode := #Status.Diagnostic.ReasonCode; END_IF;
    "FRK_PartEvent"(AlarmLog := #AlarmLog, Reason := 2027, Uid := #Part.Uid, SourcePath := #Status.Name);
    #Part.Present := FALSE;
END_FUNCTION

FUNCTION "FRK_UnitSetPermit" : Void
{ S7_Optimized_Access := 'TRUE' }
VERSION : 0.1
VAR_INPUT
    Ok : Bool;
    Diag : "ST_Diagnostic";
END_VAR
VAR_IN_OUT
    Unit : "FRK_Unit";
END_VAR
BEGIN
    #Unit.Permit := #Ok;
    #Unit.PermitDiag := #Diag;
END_FUNCTION

FUNCTION "FRK_ReleaseReason" : Void
{ S7_Optimized_Access := 'TRUE' }
VERSION : 0.1
VAR_INPUT
    Description : WString;
    Reason : DInt;
    Path : WString;
    Kind : DInt;
END_VAR
VAR_IN_OUT
    Report : "ST_ReleaseReport";
END_VAR
BEGIN
    #Report.Released := FALSE;
    IF #Report.Count < 24 THEN
        #Report.Count := #Report.Count + 1;
        #Report.Reasons[#Report.Count].Description := #Description;
        #Report.Reasons[#Report.Count].ReasonCode := #Reason;
        #Report.Reasons[#Report.Count].SourcePath := #Path;
        #Report.Reasons[#Report.Count].Kind := #Kind;
        #Report.Reasons[#Report.Count].Bypassable := FALSE;
    END_IF;
END_FUNCTION

FUNCTION "FRK_UnitOperation" : Void
{ S7_Optimized_Access := 'TRUE' }
VERSION : 0.1
VAR_INPUT
    Supported : Array[0..6] of Bool;
    Request : "ST_HmiRequest";
    Trusted : Bool;
END_VAR
VAR_IN_OUT
    Core : "FRK_Core";
    Unit : "FRK_Unit";
    Status : "ST_ModuleStatus";
    Policy : Array[0..6] of "ST_ModePolicy";
    Access : "FRK_Access";
    Response : "ST_HmiResponse";
END_VAR
VAR_TEMP
    Gate : DInt;
    Desired : DInt;
    Query : Bool;
    Level : DInt;
END_VAR
BEGIN
    #Response.Accepted := FALSE;
    #Response.Diagnostic := WSTRING#'';
    #Response.Report.Count := 0;
    #Response.Report.Released := TRUE;
    #Gate := -1;
    #Desired := -1;
    #Query := FALSE;
    CASE #Request.Kind OF
        5: #Gate := 5; #Desired := 0;
        6: #Gate := 5; #Desired := 1;
        3:
            #Gate := 4; #Desired := #Request.IntValue;
            IF #Desired = -1 THEN #Desired := -2; END_IF;
        9: #Gate := 7;
        11: #Gate := 2;
        24, 25: #Gate := 8;
        15: #Gate := 5; #Desired := 0; #Query := TRUE;
        16: #Gate := 2; #Query := TRUE;
        17: #Gate := #Request.IntValue; #Desired := -1; #Query := TRUE;
        ELSE #Gate := -1;
    END_CASE;
    IF #Gate <> -1 OR #Request.Kind = 17 THEN
        "FRK_UnitRelease"(Core := #Core, Unit := #Unit, Status := #Status, Policy := #Policy, Access := #Access, Supported := #Supported, Report := #Response.Report, Gate := #Gate, Desired := #Desired, Trusted := #Trusted);
        IF #Query THEN
            #Response.Accepted := TRUE;
        ELSIF #Response.Report.Released THEN
            CASE #Request.Kind OF
                5:
                    #Unit.StopReq := FALSE;
                    #Unit.RunReq := TRUE;
                    #Response.Accepted := TRUE;
                6:
                    #Unit.StopReq := #Core.Exec = 1;
                    IF NOT #Unit.StopReq THEN #Unit.RunReq := FALSE; END_IF;
                    #Unit.FollowStart := FALSE;
                    #Response.Accepted := TRUE;
                3:
                    IF #Desired <> #Unit.Mode THEN
                        #Unit.ExitFirst := TRUE;
                        #Unit.ModeSince := "FRK_Clock".NowMs;
                        #Unit.RequestedMode := #Desired;
                        #Unit.ModePending := TRUE;
                        IF #Unit.Mode = 1 THEN
                            #Unit.ReleaseChildren := TRUE;
                            #Unit.Clearing := TRUE;
                        END_IF;
                    END_IF;
                    #Response.Accepted := TRUE;
                9:
                    #Unit.EvReset := TRUE;
                    #Unit.ModePending := FALSE;
                    #Unit.ExitFirst := FALSE;
                    #Unit.RunReq := FALSE;
                    #Unit.AbortReq := #Core.Exec = 1;
                    #Unit.StopReq := FALSE;
                    #Unit.FollowStart := FALSE;
                    #Unit.ReleaseChildren := TRUE;
                    #Unit.Clearing := TRUE;
                    #Unit.FaultLatched := FALSE;
                    IF #Core.Exec = 3 THEN #Core.Armed := TRUE; END_IF;
                    #Response.Accepted := TRUE;
                24:
                    #Level := -1;
                    IF #Request.TextValue = WSTRING#'0' THEN #Level := 0;
                    ELSIF #Request.TextValue = WSTRING#'1' THEN #Level := 1;
                    ELSIF #Request.TextValue = WSTRING#'2' THEN #Level := 2;
                    ELSIF #Request.TextValue = WSTRING#'3' THEN #Level := 3;
                    ELSIF #Request.TextValue = WSTRING#'4' THEN #Level := 4;
                    END_IF;
                    IF #Request.IntValue >= 0 AND #Request.IntValue <= 11 AND #Level >= 0 THEN
                        IF #Request.IntValue <> 8 OR #Level <= #Access.CurrentLevel THEN
                            #Access.Policy.Required[#Request.IntValue] := #Level;
                            #Response.Accepted := TRUE;
                        END_IF;
                    END_IF;
                25:
                    IF #Request.DurationMs <= 604800000 THEN
                        #Access.Policy.SessionTimeout := DINT_TO_TIME(UDINT_TO_DINT(#Request.DurationMs));
                        #Response.Accepted := TRUE;
                    END_IF;
                ELSE
                    // Manual acceptance is resolved by the generated typed route.
                    #Response.Accepted := FALSE;
            END_CASE;
        END_IF;
    ELSE
        CASE #Request.Kind OF
            1:
                "FRK_AccessLogin"(Access := #Access, User := #Request.User, Secret := #Request.Secret, Sequence := #Request.Sequence);
                // Consumption is acknowledged now; correlated result is asynchronous.
                #Response.Accepted := TRUE;
            2:
                "FRK_AccessLogout"(Access := #Access);
                #Response.Accepted := TRUE;
            ELSE
                #Response.Diagnostic := WSTRING#'std.error.unsupportedHmiRequest';
        END_CASE;
    END_IF;
    IF #Response.Accepted AND NOT #Query THEN
        IF #Request.Kind = 5 OR #Request.Kind = 6 OR #Request.Kind = 3 OR #Request.Kind = 9 THEN
            #Unit.CascadePending := TRUE;
            #Unit.CascadeKind := #Request.Kind;
            #Unit.CascadeMode := #Unit.Mode;
            IF #Request.Kind = 3 THEN #Unit.CascadeMode := #Desired; END_IF;
        END_IF;
    END_IF;
    IF NOT #Response.Accepted AND #Request.Kind <> 11 THEN
        IF #Response.Diagnostic = WSTRING#'' THEN #Response.Diagnostic := WSTRING#'std.error.hmiRequestRejected'; END_IF;
        IF #Response.Report.Released THEN
            "FRK_ReleaseReason"(Report := #Response.Report, Description := #Response.Diagnostic, Reason := 2002, Path := STRING_TO_WSTRING(#Status.Name), Kind := 4);
        END_IF;
    END_IF;
END_FUNCTION

FUNCTION "FRK_UnitMailbox" : Void
{ S7_Optimized_Access := 'TRUE' }
VERSION : 0.1
VAR_INPUT
    Supported : Array[0..6] of Bool;
END_VAR
VAR_IN_OUT
    Core : "FRK_Core";
    Unit : "FRK_Unit";
    Status : "ST_ModuleStatus";
    Policy : Array[0..6] of "ST_ModePolicy";
    Access : "FRK_Access";
    Request : "ST_HmiRequest";
    Response : "ST_HmiResponse";
END_VAR
VAR_TEMP
    SequenceBefore : UDInt;
END_VAR
BEGIN
    #SequenceBefore := #Request.Sequence;
    IF #SequenceBefore = 0 OR #SequenceBefore = #Unit.SeenSequence THEN RETURN; END_IF;
    #Unit.Request := #Request;
    IF #Request.Sequence <> #SequenceBefore THEN #Unit.Request.Secret := ''; RETURN; END_IF;
    #Request.Secret := '';
    #Unit.RequestUser := #Access.CurrentUser;
    #Unit.SeenSequence := #SequenceBefore;
    #Unit.RequestPending := TRUE;
END_FUNCTION

FUNCTION "FRK_UnitConsume" : Void
{ S7_Optimized_Access := 'TRUE' }
VERSION : 0.1
VAR_INPUT
    Supported : Array[0..6] of Bool;
END_VAR
VAR_IN_OUT
    Core : "FRK_Core";
    Unit : "FRK_Unit";
    Status : "ST_ModuleStatus";
    Policy : Array[0..6] of "ST_ModePolicy";
    Access : "FRK_Access";
    Response : "ST_HmiResponse";
END_VAR
BEGIN
    IF NOT #Unit.RequestPending THEN RETURN; END_IF;
    // The generated typed ownership walk serves the static manifest after children.
    IF #Unit.Request.Kind = 23 THEN
        #Unit.Request.Secret := '';
        RETURN;
    END_IF;
    "FRK_UnitOperation"(Core := #Core, Unit := #Unit, Status := #Status, Policy := #Policy, Access := #Access, Supported := #Supported, Request := #Unit.Request, Response := #Response, Trusted := FALSE);
    #Unit.Request.Secret := '';
END_FUNCTION

FUNCTION "FRK_UnitMode" : Void
{ S7_Optimized_Access := 'TRUE' }
VERSION : 0.1
VAR_IN_OUT
    Core : "FRK_Core";
    Unit : "FRK_Unit";
END_VAR
BEGIN
    IF #Unit.ModePending THEN
        IF #Core.Exec = 1 THEN
            #Core.EvModeExit := TRUE;
            #Core.HookResult := 0;
        ELSIF #Core.Exec = 0 AND NOT #Unit.Clearing THEN
            #Unit.Mode := #Unit.RequestedMode;
            #Unit.ModePending := FALSE;
            #Unit.ExitFirst := FALSE;
            #Core.EvModeChanged := TRUE;
        ELSE
            #Unit.RunReq := FALSE;
        END_IF;
    END_IF;
END_FUNCTION

FUNCTION "FRK_UnitModeResolve" : Void
{ S7_Optimized_Access := 'TRUE' }
VERSION : 0.1
VAR_INPUT
    Policy : Array[0..6] of "ST_ModePolicy";
    Timeout : Time;
END_VAR
VAR_IN_OUT
    Core : "FRK_Core";
    Unit : "FRK_Unit";
    Status : "ST_ModuleStatus";
END_VAR
BEGIN
    IF #Unit.ModePending THEN
        IF #Timeout <= T#0ms OR "FRK_Elapsed"(NewMs := "FRK_Clock".NowMs, OldMs := #Unit.ModeSince) >= DINT_TO_UDINT(TIME_TO_DINT(#Timeout)) THEN
            "FRK_Fault"(Core := #Core, Status := #Status, ReasonCode := 2001, Description := WSTRING#'std.error.hmiRequestRejected');
            #Unit.ModePending := FALSE;
            #Unit.FollowStart := FALSE;
            #Unit.ReleaseChildren := TRUE;
            #Unit.Clearing := TRUE;
        ELSIF #Core.EvModeExit THEN
            #Unit.ExitFirst := FALSE;
            IF #Policy[#Unit.Mode].Style = 0 THEN
                #Unit.StopReq := TRUE;
            ELSIF #Core.HookResult <= 0 THEN
                #Unit.AbortReq := TRUE;
                #Unit.ReleaseChildren := TRUE;
                #Unit.Clearing := TRUE;
            END_IF;
        END_IF;
    END_IF;
END_FUNCTION

FUNCTION "FRK_UnitRunStart" : Void
{ S7_Optimized_Access := 'TRUE' }
VERSION : 0.1
VAR_INPUT
    Timeout : Time;
    Label : String;
END_VAR
VAR_IN_OUT
    Core : "FRK_Core";
    Status : "ST_ModuleStatus";
END_VAR
BEGIN
    "FRK_Start"(Core := #Core, Status := #Status, Supported := TRUE, Timeout := #Timeout, Label := #Label);
    // A continuous run ends at Stop. Bounded commands/steps own progress timeouts.
    #Core.TimeoutMs := 0;
END_FUNCTION

FUNCTION "FRK_DescendantsReady" : Bool
{ S7_Optimized_Access := 'TRUE' }
VERSION : 0.1
VAR_INPUT
    OwnerIndex : DInt;
END_VAR
VAR_TEMP
    Index : DInt;
    Parent : DInt;
    Depth : DInt;
END_VAR
BEGIN
    #FRK_DescendantsReady := FALSE;
    IF "FRK_Registry".Fault OR #OwnerIndex < 1 OR #OwnerIndex > "FRK_Registry".Count OR "FRK_Registry".Count > 32 THEN RETURN; END_IF;
    FOR #Index := 1 TO "FRK_Registry".Count DO
        #Parent := "FRK_Registry".Rows[#Index].Parent;
        FOR #Depth := 1 TO 32 DO
            IF #Parent = #OwnerIndex THEN
                IF "FRK_Registry".Rows[#Index].Exec <> 0 THEN RETURN; END_IF;
                EXIT;
            END_IF;
            IF #Parent = 0 THEN EXIT; END_IF;
            IF #Parent < 1 OR #Parent > "FRK_Registry".Count THEN RETURN; END_IF;
            #Parent := "FRK_Registry".Rows[#Parent].Parent;
        END_FOR;
        IF #Depth > 32 AND #Parent <> 0 THEN RETURN; END_IF;
    END_FOR;
    #FRK_DescendantsReady := TRUE;
END_FUNCTION

FUNCTION "FRK_UnitFinish" : Void
{ S7_Optimized_Access := 'TRUE' }
VERSION : 0.1
VAR_IN_OUT
    Core : "FRK_Core";
    Unit : "FRK_Unit";
    Response : "ST_HmiResponse";
    Status : "ST_ModuleStatus";
    Part : "ST_PartContext";
    AlarmLog : "FRK_AlarmLog";
    History : Array[1..16] of "ST_Diagnostic";
    Head : Int;
END_VAR
BEGIN
    IF #Core.Exec = 3 THEN
        IF NOT #Unit.EvReset THEN #Unit.FaultLatched := TRUE; END_IF;
        IF NOT #Unit.PrevError THEN
            IF #Head < 0 OR #Head >= 16 THEN #Head := 0; END_IF;
            #Head := #Head + 1;
            #History[#Head] := #Status.Diagnostic;
            "FRK_PartAborted"(Core := #Core, Unit := #Unit, Status := #Status, Part := #Part, AlarmLog := #AlarmLog);
        END_IF;
    END_IF;
    #Unit.PrevError := #Core.Exec = 3;
    IF #Core.Exec = 2 OR #Core.Exec = 4 THEN #Unit.RunReq := FALSE; END_IF;
    IF #Unit.Clearing AND #Core.Exec = 0 THEN
        IF "FRK_DescendantsReady"(OwnerIndex := #Core.RegIndex) THEN #Unit.Clearing := FALSE; END_IF;
    END_IF;
    #Unit.AbortReq := FALSE;
    #Unit.ReleaseChildren := FALSE;
    #Unit.EvReset := FALSE;
    IF #Unit.RequestPending THEN
        #Response.AckSequence := #Unit.SeenSequence;
        #Unit.RequestPending := FALSE;
    END_IF;
END_FUNCTION

// Shared Unit routing: typed generated edges carry these owning predicates.
FUNCTION "FRK_PathOwned" : Bool
{ S7_Optimized_Access := 'TRUE' }
VERSION : 0.1
VAR_INPUT
    OwnerPath : String;
    TargetPath : WString;
END_VAR
VAR_TEMP
    Width : Int;
END_VAR
BEGIN
    #FRK_PathOwned := FALSE;
    #Width := LEN(#OwnerPath);
    IF #Width = 0 THEN RETURN; END_IF;
    IF #TargetPath = STRING_TO_WSTRING(#OwnerPath) THEN #FRK_PathOwned := TRUE; RETURN; END_IF;
    IF LEN(#TargetPath) <= #Width THEN RETURN; END_IF;
    #FRK_PathOwned := LEFT(IN := #TargetPath, L := #Width) = STRING_TO_WSTRING(#OwnerPath) AND #TargetPath[#Width + 1] = WCHAR#'.';
END_FUNCTION

FUNCTION "FRK_UnitRelease" : Void
{ S7_Optimized_Access := 'TRUE' }
VERSION : 0.1
VAR_INPUT
    Gate : DInt;
    Desired : DInt;
    Trusted : Bool;
    Core : "FRK_Core";
    Unit : "FRK_Unit";
    Status : "ST_ModuleStatus";
    Policy : Array[0..6] of "ST_ModePolicy";
    Access : "FRK_Access";
    Supported : Array[0..6] of Bool;
END_VAR
VAR_IN_OUT
    Report : "ST_ReleaseReport";
END_VAR
BEGIN
    #Report.Count := 0;
    #Report.Released := TRUE;
    IF #Gate <> 5 AND #Gate <> 4
        AND #Gate <> 7 AND #Gate <> 2
        AND #Gate <> 8
        AND NOT (#Unit.ConfigEnabled AND #Gate = 1)
        AND NOT (#Unit.ModelEnabled AND #Gate = 3) THEN
        "FRK_ReleaseReason"(Report := #Report, Description := WSTRING#'std.error.unsupportedHmiRequest', Reason := 2008, Path := STRING_TO_WSTRING(#Status.Name), Kind := 4);
        RETURN;
    END_IF;
    IF NOT #Trusted THEN
        IF #Access.CurrentLevel < #Access.Policy.Required[#Gate] THEN
            "FRK_ReleaseReason"(Report := #Report, Description := WSTRING#'std.release.insufficientAction', Reason := 2002, Path := STRING_TO_WSTRING(#Status.Name), Kind := 1);
        END_IF;
    END_IF;
    CASE #Gate OF
        3:
            IF #Core.Exec <> 0 OR #Unit.ModePending OR #Unit.Clearing OR NOT "FRK_DescendantsReady"(OwnerIndex := #Core.RegIndex) THEN
                "FRK_ReleaseReason"(Report := #Report, Description := WSTRING#'std.error.hmiRequestRejected', Reason := 2011, Path := STRING_TO_WSTRING(#Status.Name), Kind := 4);
            END_IF;
            IF #Unit.AlarmBlocking THEN
                "FRK_ReleaseReason"(Report := #Report, Description := WSTRING#'std.release.manualReset', Reason := 0, Path := STRING_TO_WSTRING(#Status.Name), Kind := 2);
            END_IF;
            IF NOT #Unit.Permit THEN
                "FRK_ReleaseReason"(Report := #Report, Description := #Unit.PermitDiag.Description, Reason := #Unit.PermitDiag.ReasonCode, Path := #Unit.PermitDiag.SourcePath, Kind := 3);
            END_IF;
        5:
            // Desired=0 is Start, Desired=1 is Stop. Generic action query is Stop.
            IF #Desired = 0 THEN
                IF #Unit.Mode = 1 OR #Unit.ModePending THEN
                    "FRK_ReleaseReason"(Report := #Report, Description := WSTRING#'std.error.unsupportedModeRequest', Reason := 2002, Path := STRING_TO_WSTRING(#Status.Name), Kind := 0);
                END_IF;
                IF #Core.Exec <> 0 OR #Unit.RunReq OR #Unit.Clearing OR #Unit.FaultLatched THEN
                    "FRK_ReleaseReason"(Report := #Report, Description := WSTRING#'std.error.hmiRequestRejected', Reason := 2011, Path := STRING_TO_WSTRING(#Status.Name), Kind := 4);
                END_IF;
                IF #Unit.AlarmBlocking THEN
                    "FRK_ReleaseReason"(Report := #Report, Description := WSTRING#'std.release.manualReset', Reason := 0, Path := STRING_TO_WSTRING(#Status.Name), Kind := 2);
                END_IF;
                IF #Unit.ConfigBlocked THEN
                    "FRK_ReleaseReason"(Report := #Report, Description := WSTRING#'std.release.configRestoreUnacknowledged', Reason := 2040, Path := STRING_TO_WSTRING(#Status.Name), Kind := 2);
                END_IF;
                IF NOT #Unit.Permit THEN
                    "FRK_ReleaseReason"(Report := #Report, Description := #Unit.PermitDiag.Description, Reason := #Unit.PermitDiag.ReasonCode, Path := #Unit.PermitDiag.SourcePath, Kind := 3);
                END_IF;
            END_IF;
        4:
            IF #Unit.ModePending THEN
                "FRK_ReleaseReason"(Report := #Report, Description := WSTRING#'std.release.modeChangeAlreadyPending', Reason := 2011, Path := STRING_TO_WSTRING(#Status.Name), Kind := 0);
            END_IF;
            IF #Core.Exec = 1 AND #Unit.Mode <> 1 THEN
                IF #Policy[#Unit.Mode].Shield = 2 THEN
                    "FRK_ReleaseReason"(Report := #Report, Description := WSTRING#'std.release.modeSwitchBlockedWhileRunning', Reason := 2002, Path := STRING_TO_WSTRING(#Status.Name), Kind := 0);
                END_IF;
            END_IF;
            IF #Desired <> -1 THEN
                IF #Desired < 0 OR #Desired >= 7 THEN
                    "FRK_ReleaseReason"(Report := #Report, Description := WSTRING#'std.error.unsupportedModeRequest', Reason := 2008, Path := STRING_TO_WSTRING(#Status.Name), Kind := 0);
                ELSIF NOT #Supported[#Desired] THEN
                    "FRK_ReleaseReason"(Report := #Report, Description := WSTRING#'std.error.unsupportedModeRequest', Reason := 2008, Path := STRING_TO_WSTRING(#Status.Name), Kind := 0);
                END_IF;
            END_IF;
        7:
            // The complete alarm model is separate; this gate owns the current latch.
            IF NOT #Unit.FaultLatched AND NOT #Unit.AlarmBlocking AND #Core.Exec = 0 AND NOT #Unit.Clearing AND NOT #Unit.ModePending AND NOT #Unit.FollowStart THEN
                IF "FRK_DescendantsReady"(OwnerIndex := #Core.RegIndex) THEN
                    "FRK_ReleaseReason"(Report := #Report, Description := WSTRING#'std.release.noBlockingAlarm', Reason := 2011, Path := STRING_TO_WSTRING(#Status.Name), Kind := 4);
                END_IF;
            END_IF;
        2:
            "FRK_ManualCommon"(Core := #Core, Unit := #Unit, Status := #Status, Report := #Report);
        ELSE
            RETURN;
    END_CASE;
END_FUNCTION

FUNCTION "FRK_ManualCommon" : Void
{ S7_Optimized_Access := 'TRUE' }
VERSION : 0.1
VAR_INPUT
    Core : "FRK_Core";
    Unit : "FRK_Unit";
    Status : "ST_ModuleStatus";
END_VAR
VAR_IN_OUT
    Report : "ST_ReleaseReport";
END_VAR
BEGIN
    IF #Unit.Mode <> 1 OR #Unit.ModePending THEN
        "FRK_ReleaseReason"(Report := #Report, Description := WSTRING#'std.release.manualModeRequired', Reason := 2002, Path := STRING_TO_WSTRING(#Status.Name), Kind := 0);
    END_IF;
    IF #Core.Exec <> 0 OR #Unit.Clearing OR #Unit.FaultLatched THEN
        "FRK_ReleaseReason"(Report := #Report, Description := WSTRING#'std.error.hmiRequestRejected', Reason := 2011, Path := STRING_TO_WSTRING(#Status.Name), Kind := 4);
    END_IF;
    IF #Unit.AlarmBlocking THEN
        "FRK_ReleaseReason"(Report := #Report, Description := WSTRING#'std.release.manualReset', Reason := 0, Path := STRING_TO_WSTRING(#Status.Name), Kind := 2);
    END_IF;
    IF NOT #Unit.Permit THEN
        "FRK_ReleaseReason"(Report := #Report, Description := #Unit.PermitDiag.Description, Reason := #Unit.PermitDiag.ReasonCode, Path := #Unit.PermitDiag.SourcePath, Kind := 3);
    END_IF;
END_FUNCTION

FUNCTION "FRK_ManualCondition" : Void
{ S7_Optimized_Access := 'TRUE' }
VERSION : 0.1
VAR_INPUT
    Slot : Int;
    Value : DInt;
    Ok : Bool;
    Diag : "ST_Diagnostic";
    Bypassable : Bool;
END_VAR
VAR_IN_OUT
    Conditions : Array[1..16] of "FRK_ManualConditionRow";
END_VAR
BEGIN
    IF #Slot < 1 OR #Slot > 16 THEN RETURN; END_IF;
    #Conditions[#Slot].Used := TRUE;
    #Conditions[#Slot].Value := #Value;
    #Conditions[#Slot].Ok := #Ok;
    #Conditions[#Slot].Diag := #Diag;
    #Conditions[#Slot].Bypassable := #Bypassable;
END_FUNCTION

FUNCTION "FRK_ManualApply" : Void
{ S7_Optimized_Access := 'TRUE' }
VERSION : 0.1
VAR_INPUT
    Request : "ST_HmiRequest";
    Status : "ST_ModuleStatus";
    Core : "FRK_Core";
    Commands : Array[1..12] of "ST_CommandInfo";
    Count : DInt;
    Conditions : Array[1..16] of "FRK_ManualConditionRow";
END_VAR
VAR_IN_OUT
    Report : "ST_ReleaseReport";
    Execute : Bool;
    Command : DInt;
    ManualOwned : Bool;
END_VAR
VAR_TEMP
    Index : Int;
    Supported : Bool;
    PreviousCount : Int;
END_VAR
BEGIN
    #Supported := FALSE;
    IF #Count >= 0 AND #Count <= 12 THEN
        FOR #Index := 1 TO DINT_TO_INT(#Count) DO
            IF #Commands[#Index].Value = #Request.IntValue AND #Commands[#Index].Style = 0 THEN #Supported := TRUE; END_IF;
        END_FOR;
    END_IF;
    IF NOT #Supported THEN
        "FRK_ReleaseReason"(Report := #Report, Description := WSTRING#'std.error.unsupportedHmiRequest', Reason := 2008, Path := STRING_TO_WSTRING(#Status.Name), Kind := 4);
    END_IF;
    IF #Core.Exec <> 0 OR #Execute OR #Core.ReleasePending THEN
        "FRK_ReleaseReason"(Report := #Report, Description := WSTRING#'std.error.hmiRequestRejected', Reason := 2011, Path := STRING_TO_WSTRING(#Status.Name), Kind := 4);
    END_IF;
    FOR #Index := 1 TO 16 DO
        IF #Conditions[#Index].Used AND NOT #Conditions[#Index].Ok THEN
            IF #Conditions[#Index].Value = 0 OR #Conditions[#Index].Value = #Request.IntValue THEN
                #PreviousCount := #Report.Count;
                "FRK_ReleaseReason"(Report := #Report, Description := #Conditions[#Index].Diag.Description, Reason := #Conditions[#Index].Diag.ReasonCode, Path := STRING_TO_WSTRING(#Status.Name), Kind := 3);
                IF #Report.Count > #PreviousCount THEN #Report.Reasons[#Report.Count].Bypassable := #Conditions[#Index].Bypassable; END_IF;
            END_IF;
        END_IF;
    END_FOR;
    IF #Request.Kind = 11 AND #Report.Released THEN
        #Command := #Request.IntValue;
        #Execute := TRUE;
        #ManualOwned := TRUE;
    END_IF;
END_FUNCTION

FUNCTION "FRK_ManualFinish" : Void
{ S7_Optimized_Access := 'TRUE' }
VERSION : 0.1
VAR_INPUT
    Core : "FRK_Core";
END_VAR
VAR_IN_OUT
    Execute : Bool;
    ManualOwned : Bool;
END_VAR
BEGIN
    IF #ManualOwned AND #Core.Exec <> 1 THEN
        #Execute := FALSE;
        #ManualOwned := FALSE;
    END_IF;
END_FUNCTION

FUNCTION "FRK_UnitCascade" : Void
{ S7_Optimized_Access := 'TRUE' }
VERSION : 0.1
VAR_INPUT
    ParentUnit : "FRK_Unit";
    Supported : Array[0..6] of Bool;
END_VAR
VAR_IN_OUT
    Core : "FRK_Core";
    Unit : "FRK_Unit";
    Status : "ST_ModuleStatus";
    Policy : Array[0..6] of "ST_ModePolicy";
    Access : "FRK_Access";
    AlarmLog : "FRK_AlarmLog";
END_VAR
VAR_TEMP
    Request : "ST_HmiRequest";
END_VAR
BEGIN
    IF NOT #ParentUnit.CascadePending THEN RETURN; END_IF;
    IF #ParentUnit.CascadeKind = 6 OR #ParentUnit.CascadeKind = 9 THEN
        #Unit.FollowStart := FALSE;
        #Request.Kind := #ParentUnit.CascadeKind;
        "FRK_UnitOperation"(Core := #Core, Unit := #Unit, Status := #Status, Policy := #Policy, Access := #Access, Supported := #Supported, Request := #Request, Response := "FRK_UnitScratch".Response, Trusted := TRUE);
        RETURN;
    END_IF;
    #Request.Kind := 3;
    #Request.IntValue := #ParentUnit.CascadeMode;
    "FRK_UnitOperation"(Core := #Core, Unit := #Unit, Status := #Status, Policy := #Policy, Access := #Access, Supported := #Supported, Request := #Request, Response := "FRK_UnitScratch".Response, Trusted := TRUE);
    IF NOT "FRK_UnitScratch".Response.Accepted THEN
        #Unit.FollowStart := FALSE;
        #Request.Kind := 6;
        "FRK_UnitOperation"(Core := #Core, Unit := #Unit, Status := #Status, Policy := #Policy, Access := #Access, Supported := #Supported, Request := #Request, Response := "FRK_UnitScratch".Response, Trusted := TRUE);
        // Core names this event but has no assigned E_Reason ordinal yet.
        "FRK_AlarmMessage"(AlarmLog := #AlarmLog, Reason := 2008, Description := WSTRING#'std.event.childModeUnsupported', SourcePath := STRING_TO_WSTRING(#Status.Name));
    ELSE
        #Unit.FollowStart := #ParentUnit.CascadeKind = 5;
    END_IF;
END_FUNCTION

FUNCTION "FRK_UnitFollow" : Void
{ S7_Optimized_Access := 'TRUE' }
VERSION : 0.1
VAR_INPUT
    Supported : Array[0..6] of Bool;
END_VAR
VAR_IN_OUT
    Core : "FRK_Core";
    Unit : "FRK_Unit";
    Status : "ST_ModuleStatus";
    Policy : Array[0..6] of "ST_ModePolicy";
    Access : "FRK_Access";
END_VAR
VAR_TEMP
    Request : "ST_HmiRequest";
END_VAR
BEGIN
    IF #Unit.FollowStart AND NOT #Unit.ModePending AND NOT #Unit.Clearing THEN
        #Unit.FollowStart := FALSE;
        #Request.Kind := 5;
        "FRK_UnitOperation"(Core := #Core, Unit := #Unit, Status := #Status, Policy := #Policy, Access := #Access, Supported := #Supported, Request := #Request, Response := "FRK_UnitScratch".Response, Trusted := TRUE);
    END_IF;
END_FUNCTION
